Fanuc KAREL source: kt00489.KL

-- PROVISIONAL review KL for V770-1; original PC SHA256 b87e1a059f767ca21b8d9d8c8d08725f8356ab26509ccbf1067e98c2783f8764
-- Incomplete behavior may be omitted. Consult companion uncertainty JSON. Do not deploy.
PROGRAM KT00489
%NOLOCKGROUP
-- UNRESOLVED_DECL P1 type=000101
-- UNRESOLVED_DECL P2 type=000199
-- UNRESOLVED_DECL OUT type=000101
BEGIN
  -- UNRESOLVED_PC offsets 5-34; opcodes 49,49,7E,60,4A
  -- UNRESOLVED_PC offsets 39-43; opcodes 7F
END KT00489
